(* IEC 61131-3 sources: rusty/tests/lit/single/property, 21 files *)

(* ---- called_inside_pou_where_defined.st ---- *)
// RUN: %COMPILE %s && %RUN | %CHECK %s

FUNCTION_BLOCK A
    PROPERTY_GET sayCheese: DINT
        printf('Cheese');
    END_PROPERTY

    sayCheese;
END_FUNCTION_BLOCK

FUNCTION main
    VAR
        instanceA : A;
    END_VAR

    // CHECK: Cheese
    instanceA();
END_FUNCTION

(* ---- complex.st ---- *)
// RUN: %COMPILE %s && %RUN | %CHECK %s
FUNCTION_BLOCK fb
VAR
  x : DINT;
  foo: nest_level1;
  END_VAR
END_FUNCTION_BLOCK

FUNCTION_BLOCK nest_level1
VAR
  foo: nest_level2;
END_VAR
END_FUNCTION_BLOCK

FUNCTION_BLOCK nest_level2
VAR
  foo: DINT := 0;
END_VAR
    PROPERTY_GET myProp: DINT
      myProp := foo + 5;
    END_PROPERTY

    PROPERTY_SET myProp: DINT
      foo := myProp + foo;
    END_PROPERTY
END_FUNCTION_BLOCK

FUNCTION main
    VAR
        bar: fb;
        x : DINT := 1;
    END_VAR

printf('%d$N', bar.foo.foo.myProp);   // CHECK: 5
bar.foo.foo.myProp := 10;
printf('%d$N', bar.foo.foo.myProp);   // CHECK: 15
END_FUNCTION

(* ---- get_with_early_return.st ---- *)
// RUN: %COMPILE %s && %RUN | %CHECK %s

// A RETURN in a getter returns the value of the property variable at the RETURN
FUNCTION_BLOCK fb
    VAR_INPUT
        mode : DINT;
    END_VAR

    PROPERTY_GET p : DINT
        IF mode = 1 THEN
            p := 5;
            RETURN;
        END_IF

        CASE mode OF
            2:
                p := 7;
                RETURN;
        END_CASE

        WHILE TRUE DO
            p := 8;
            IF mode = 3 THEN
                RETURN;
            END_IF
            EXIT;
        END_WHILE

        p := 6;
    END_PROPERTY
END_FUNCTION_BLOCK

FUNCTION main : DINT
    VAR
        f : fb;
    END_VAR

    // CHECK: 6
    printf('%d$N', f.p);

    f.mode := 1;
    // CHECK: 5
    printf('%d$N', f.p);

    f.mode := 2;
    // CHECK: 7
    printf('%d$N', f.p);

    f.mode := 3;
    // CHECK: 8
    printf('%d$N', f.p);
END_FUNCTION

(* ---- getter_used_in_array_indexing.st ---- *)
// RUN: %COMPILE %s && %RUN | %CHECK %s

FUNCTION_BLOCK fb
    VAR
        localVariable: ARRAY[1..5] OF DINT := [2, 4, 8, 16, 32];
    END_VAR

    PROPERTY_GET foo: ARRAY[1..5] OF DINT
        foo := localVariable;
    END_PROPERTY

    PROPERTY_GET bar: DINT
        bar := 3;
    END_PROPERTY
END_FUNCTION_BLOCK

FUNCTION main
    VAR
        instance: fb;

        arrayValue: ARRAY[1..5] OF DINT;
        arrayIndex: DINT;
    END_VAR

    printf('%d$N', instance.foo[instance.bar]); // CHECK: 8
END_FUNCTION

(* ---- modify_array_value_with_get_and_set.st ---- *)
// RUN: %COMPILE %s && %RUN | %CHECK %s

FUNCTION_BLOCK fb
    VAR
        localArray: ARRAY[1..5] OF DINT := [1, 2, 3, 4, 5];
    END_VAR

    PROPERTY_GET foo: ARRAY[1..5] OF DINT
        foo := localArray;
    END_PROPERTY

    PROPERTY_SET foo: ARRAY[1..5] OF DINT
        localArray := foo;
    END_PROPERTY
END_FUNCTION_BLOCK

FUNCTION main
    VAR
        localArray: ARRAY[1..5] OF DINT;
        fbInstance: fb;
    END_VAR

    localArray := fbInstance.foo;
    localArray[1] := 5;
    localArray[5] := 1;

    fbInstance.foo := localArray;

    printf('%d$N', fbInstance.foo[1]); // CHECK: 5
    printf('%d$N', fbInstance.foo[5]); // CHECK: 1
END_FUNCTION

(* ---- multiply_properties_single_pou.st ---- *)
// RUN: %COMPILE %s && %RUN | %CHECK %s

FUNCTION_BLOCK A
    VAR
        foo : DINT;
    END_VAR

    PROPERTY_GET increaseFooBy10: DINT
        printf('Inside increaseFooBy10$N');
        foo := foo + 10;
    END_PROPERTY

    PROPERTY_GET increaseFooBy20: DINT
        printf('Inside increaseFooBy20$N');
        foo := foo + 20;
    END_PROPERTY

    PROPERTY_GET increaseFooBy30: DINT
        printf('Inside increaseFooBy30$N');
        increaseFooBy20;
        increaseFooBy10;
    END_PROPERTY

    PROPERTY_GET readFoo: DINT
        printf('Inside readFoo$N');
        readFoo := foo;
    END_PROPERTY
END_FUNCTION_BLOCK

FUNCTION main
    VAR
        instanceA : A;
        result : DINT;
    END_VAR

    // CHECK: Inside increaseFooBy10
    instanceA.increaseFooBy10;

    // CHECK: Inside increaseFooBy20
    instanceA.increaseFooBy20;

    // CHECK: Inside increaseFooBy30
    // CHECK: Inside increaseFooBy20
    // CHECK: Inside increaseFooBy10
    instanceA.increaseFooBy30;

    // CHECK: Inside readFoo
    // CHECK: 60
    printf('%d$N', instanceA.readFoo);
END_FUNCTION

(* ---- nested.st ---- *)
// RUN: %COMPILE %s && %RUN | %CHECK %s

FUNCTION_BLOCK A
    VAR
        instanceB : B;
    END_VAR
END_FUNCTION_BLOCK

FUNCTION_BLOCK B
    VAR
        instanceC : C;
    END_VAR
END_FUNCTION_BLOCK

FUNCTION_BLOCK C
    VAR
        localPrivateVariable : DINT := 69;
    END_VAR

    PROPERTY_GET foo: DINT
        printf('Inside getter$N');
        foo := localPrivateVariable;
    END_PROPERTY

    PROPERTY_SET foo: DINT
        printf('Inside setter$N');
        localPrivateVariable := localPrivateVariable + foo;
    END_PROPERTY
END_FUNCTION_BLOCK

FUNCTION main
    VAR
        instanceA : A;
    END_VAR

    // CHECK: Inside getter
    // CHECK: 69
    printf('%d$N', instanceA.instanceB.instanceC.foo);

    // CHECK: Inside setter
    instanceA.instanceB.instanceC.foo := 351;

    // CHECK: Inside getter
    // CHECK: 420
    printf('%d$N', instanceA.instanceB.instanceC.foo);
END_FUNCTION

(* ---- oop_extended_fb_calls_property_in_another_property.st ---- *)
// RUN: %COMPILE %s && %RUN | %CHECK %s

FUNCTION_BLOCK fb
    PROPERTY_GET foo: DINT
        foo := 69;
    END_PROPERTY
END_FUNCTION_BLOCK

FUNCTION_BLOCK fb2 EXTENDS fb
    PROPERTY_GET bar: DINT
        bar := foo;
    END_PROPERTY
END_FUNCTION_BLOCK

FUNCTION main
    VAR
        fbInstance: fb2;
    END_VAR

    printf('%d$N', fbInstance.bar); // CHECK: 69
END_FUNCTION

(* ---- oop_extended_function_block.st ---- *)
// RUN: %COMPILE %s && %RUN | %CHECK %s

FUNCTION_BLOCK fb
    VAR
        returnValue: ARRAY[1..5] OF STRING := ['a', 'b', 'c', 'd', 'e'];
    END_VAR

    PROPERTY_GET foo: ARRAY[1..5] OF STRING
        foo := returnValue;
    END_PROPERTY

    PROPERTY_GET bar: DINT
        bar := 5;
    END_PROPERTY
END_FUNCTION_BLOCK

FUNCTION_BLOCK fb2 EXTENDS fb
END_FUNCTION_BLOCK

FUNCTION main
    VAR
        fbInstance: fb2;
    END_VAR

    printf('%s$N', REF(fbInstance.foo[1])); // CHECK: a
    printf('%d$N', fbInstance.bar); // CHECK: 5
END_FUNCTION

(* ---- oop_inheritance.st ---- *)
// RUN: %COMPILE %s && %RUN | %CHECK %s

INTERFACE intf
    PROPERTY_GET prop: DINT END_PROPERTY
    PROPERTY_SET prop: DINT END_PROPERTY
END_INTERFACE

FUNCTION_BLOCK fb IMPLEMENTS intf
    VAR
        localPrivateVariable: DINT := 69;
    END_VAR

    PROPERTY_GET prop: DINT
        prop := localPrivateVariable;
    END_PROPERTY

    PROPERTY_SET prop: DINT
        // This should never be called when using fb2 because it will be overridden
        localPrivateVariable := 0;
    END_PROPERTY
END_FUNCTION_BLOCK

FUNCTION_BLOCK fb2 EXTENDS fb
    PROPERTY_SET prop: DINT
        localPrivateVariable := prop;
    END_PROPERTY
END_FUNCTION_BLOCK

FUNCTION main: DINT
    VAR
        instance: fb2;
    END_VAR

    // This will call the getter from fb
    printf('%d$N', instance.prop); // CHECK: 69

    // This will call the setter from fb2
    instance.prop := 420;
    printf('%d$N', instance.prop); // CHECK: 420
END_FUNCTION

(* ---- oop_interface_extension.st ---- *)
// RUN: %COMPILE %s && %RUN | %CHECK %s

FUNCTION_BLOCK fb1
    VAR
        localPrivateVariable: DINT := 68;
    END_VAR

    PROPERTY_GET prop: DINT
        prop := localPrivateVariable;
    END_PROPERTY
END_FUNCTION_BLOCK

FUNCTION_BLOCK fb2 EXTENDS fb1
    PROPERTY_SET prop: DINT
        VAR
            x: DINT;
        END_VAR

        x := prop + 1;
        localPrivateVariable := x;
    END_PROPERTY
END_FUNCTION_BLOCK

FUNCTION main
    VAR
        instance: fb2;
    END_VAR

    instance.prop := 68;
    printf('%d$N', instance.prop); // CHECK: 69
END_FUNCTION

(* ---- oop_interface_extension_call_in_fb_body.st ---- *)
// RUN: %COMPILE %s && %RUN | %CHECK %s

FUNCTION_BLOCK fb1
    VAR
        localPrivateVariable: DINT := 67;
    END_VAR

    PROPERTY_GET prop: DINT
        prop := localPrivateVariable;
    END_PROPERTY
END_FUNCTION_BLOCK

FUNCTION_BLOCK fb2 EXTENDS fb1
    PROPERTY_SET prop: DINT
        VAR
            x: DINT;
        END_VAR

        x := prop + 1;
        localPrivateVariable := x;
    END_PROPERTY

    prop := prop + 1;
END_FUNCTION_BLOCK

FUNCTION main
    VAR
        instance: fb2;
    END_VAR

    instance();
    printf('%d$N', instance.prop); // CHECK: 69
END_FUNCTION

(* ---- property_get_with_reference_to_return_type.st ---- *)
// RUN: %COMPILE %s && %RUN | %CHECK %s
PROGRAM test
VAR
	fb	: fb;
END_VAR

printf('%d$N', fb.myStructuredVar.x);

END_PROGRAM

FUNCTION_BLOCK fb
VAR
	_myStructuredVar	: structuredTypeOrFb;
END_VAR

PROPERTY_GET myStructuredVar : REFERENCE TO structuredTypeOrFb
	myStructuredVar REF= _myStructuredVar;
END_PROPERTY

END_FUNCTION_BLOCK

TYPE structuredTypeOrFb :
	STRUCT
		x	: INT := 42;
	END_STRUCT
END_TYPE

FUNCTION main
    // CHECK: 42
    test();
END_FUNCTION

(* ---- property_get_with_referenceto_return_type_in_expression.st ---- *)
// RUN: %COMPILE %s && %RUN | %CHECK %s
PROGRAM test
VAR
	fb : fb;
    tempStruct_store : structuredTypeOrFb;
    tempStruct : REFERENCE TO structuredTypeOrFb;
    y: INT;
END_VAR

tempStruct_store.x := 51;
tempStruct REF= tempStruct_store;

// CHECK: Pre-init value: 51
printf('Pre-init value: %d$N', tempStruct.x);

fb.myStructuredVar := tempStruct;

// CHECK: Post-init value: 51
printf('Post-init value: %d$N', fb.myStructuredVar.x);

// CHECK: Expression value: 52
y := fb.myStructuredVar.x + 1;
printf('Expression value: %d$N', y);

END_PROGRAM

FUNCTION_BLOCK fb
VAR
	_myStructuredVar	: structuredTypeOrFb;
END_VAR

PROPERTY_GET myStructuredVar : REFERENCE TO structuredTypeOrFb
	myStructuredVar REF= _myStructuredVar;
END_PROPERTY

PROPERTY_SET myStructuredVar : REFERENCE TO structuredTypeOrFb
	_myStructuredVar := myStructuredVar;
END_PROPERTY

END_FUNCTION_BLOCK

TYPE structuredTypeOrFb :
	STRUCT
		x	: INT := 42;
	END_STRUCT
END_TYPE

FUNCTION main
    test();
END_FUNCTION

(* ---- property_set_with_reference_to_return_type.st ---- *)
// RUN: %COMPILE %s && %RUN | %CHECK %s
PROGRAM test
VAR
	fb : fb;
    tempStruct_store : structuredTypeOrFb;
    tempStruct : REFERENCE TO structuredTypeOrFb;
END_VAR

tempStruct_store.x := 51;
tempStruct REF= tempStruct_store;

// CHECK: Pre-init value: 51
printf('Pre-init value: %d$N', tempStruct.x);

fb.myStructuredVar := tempStruct;

// CHECK: Post-init value: 51
printf('Post-init value: %d$N', fb.myStructuredVar.x);

END_PROGRAM

FUNCTION_BLOCK fb
VAR
	_myStructuredVar	: structuredTypeOrFb;
END_VAR

PROPERTY_GET myStructuredVar : REFERENCE TO structuredTypeOrFb
	myStructuredVar REF= _myStructuredVar;
END_PROPERTY

PROPERTY_SET myStructuredVar : REFERENCE TO structuredTypeOrFb
	_myStructuredVar := myStructuredVar;
END_PROPERTY

END_FUNCTION_BLOCK

TYPE structuredTypeOrFb :
	STRUCT
		x	: INT := 42;
	END_STRUCT
END_TYPE

FUNCTION main
    test();
END_FUNCTION

(* ---- property_used_in_action.st ---- *)
// RUN: %COMPILE %s && %RUN | %CHECK %s
FUNCTION_BLOCK A
    VAR
        x : DINT := 42;
    END_VAR
    PROPERTY_GET foo: DINT
        foo := x;
    END_PROPERTY

    METHOD bar : DINT
        bar := foo;
    END_METHOD
END_FUNCTION_BLOCK

ACTIONS
    ACTION baz
        // CHECK: 42
        printf('%d$N', bar());
        // CHECK: 42
        printf('%d$N', foo);
    END_ACTION
END_ACTIONS

FUNCTION main
    VAR
        instanceA : A;
    END_VAR
        instanceA.baz();
END_FUNCTION

(* ---- property_with_chained_reference_to_return_type.st ---- *)
// RUN: %COMPILE %s && %RUN | %CHECK %s
PROGRAM test
VAR
	fb : fb;
    y : INT;
    tempStruct_store : structuredTypeOrFb;
    tempStruct2_store : structuredTypeOrFb2;
    tempStruct : REFERENCE TO structuredTypeOrFb;
END_VAR

tempStruct2_store.x := 51;
tempStruct_store.subType REF= tempStruct2_store;
tempStruct REF= tempStruct_store;

// CHECK: Pre-init value: 51
printf('Pre-init value: %d$N', tempStruct.subType.x);

fb.myStructuredVar := tempStruct;

// CHECK: Post-init value: 51
printf('Post-init value: %d$N', fb.myStructuredVar.subType.x);

END_PROGRAM

FUNCTION_BLOCK fb
VAR
	_myStructuredVar	: structuredTypeOrFb;
END_VAR

PROPERTY_GET myStructuredVar : REFERENCE TO structuredTypeOrFb
	myStructuredVar REF= _myStructuredVar;
END_PROPERTY

PROPERTY_SET myStructuredVar : REFERENCE TO structuredTypeOrFb
	_myStructuredVar := myStructuredVar;
END_PROPERTY

END_FUNCTION_BLOCK

TYPE structuredTypeOrFb :
	STRUCT
		subType : REFERENCE TO structuredTypeOrFb2;
	END_STRUCT
END_TYPE

TYPE structuredTypeOrFb2 :
	STRUCT
		x : INT := 42;
	END_STRUCT
END_TYPE

FUNCTION main
    test();
END_FUNCTION

(* ---- property_with_local_variables.st ---- *)
// RUN: %COMPILE %s && %RUN | %CHECK %s
FUNCTION_BLOCK fb
    VAR
        localPrivateVariable: DINT := 5;
    END_VAR

    PROPERTY_GET foo: DINT
        VAR
            one: DINT := 1;
        END_VAR

        foo := localPrivateVariable + one;
    END_PROPERTY

    PROPERTY_SET foo: DINT
        VAR
            two: DINT := 2;
            three: DINT := 3;
        END_VAR
        localPrivateVariable := two + foo + three;
    END_PROPERTY
END_FUNCTION_BLOCK

FUNCTION main
    VAR
        localVariable: DINT;
        instance: fb;
    END_VAR

    // Retrieving the getter return value using another variable
    localVariable := instance.foo;
    printf('%d$N', localVariable); // CHECK: 6

    // Retrieving the getter return value using the property directly
    printf('%d$N', instance.foo); // CHECK: 6

    instance.foo := 10;
    printf('%d$N', instance.foo); // CHECK: 16
END_FUNCTION

(* ---- same_property_in_different_pous_called_in_method.st ---- *)
// RUN: %COMPILE %s && %RUN | %CHECK %s
FUNCTION_BLOCK A
    VAR
        x : DINT := 42;
    END_VAR

    PROPERTY_GET foo: DINT
        foo := x;
    END_PROPERTY
END_FUNCTION_BLOCK

FUNCTION_BLOCK B
    VAR
        x : DINT := 69;
    END_VAR

    PROPERTY_GET foo: DINT
        foo := x;
    END_PROPERTY

    METHOD bar : DINT
    VAR
        instanceA : A;
    END_VAR
        bar := foo;
    END_METHOD

    METHOD baz : DINT
    VAR
        instanceA : A;
    END_VAR
        baz := instanceA.foo;
    END_METHOD
END_FUNCTION_BLOCK

FUNCTION main
    VAR
        instanceB : B;
    END_VAR

    printf('%d$N', instanceB.bar()); // CHECK: 69
    printf('%d$N', instanceB.baz()); // CHECK: 42
END_FUNCTION

(* ---- simple.st ---- *)
// RUN: %COMPILE %s && %RUN | %CHECK %s
FUNCTION_BLOCK fb
    VAR
        localPrivateVariable : DINT := 5;
    END_VAR

    PROPERTY_GET foo: DINT
        foo := localPrivateVariable;
    END_PROPERTY

    PROPERTY_SET foo: DINT
        localPrivateVariable := foo + 5;
    END_PROPERTY
END_FUNCTION_BLOCK

FUNCTION main
    VAR
        localVariable : DINT;
        instance : fb;
    END_VAR

    // Retrieving the getter return value using another variable
    localVariable := instance.foo;
    printf('%d$N', localVariable);  // CHECK: 5

    // Retrieving the getter return value using the property directly
    printf('%d$N', instance.foo);   // CHECK: 5

    instance.foo := 10;
    printf('%d$N', instance.foo);   // CHECK: 15
END_FUNCTION

(* ---- struct_return_type.st ---- *)
// RUN: %COMPILE %s && %RUN | %CHECK %s

TYPE
    Transaction: STRUCT
        id: DINT;
        values: ARRAY[1..10] OF DINT;
    END_STRUCT
END_TYPE

FUNCTION print_txn
    VAR_INPUT {ref}
        value: Transaction;
    END_VAR

    VAR
        idx: DINT;
    END_VAR

    printf('{ id: %d, values: [', value.id);
    FOR idx := 1 TO 10 DO
        IF idx > 1 THEN
            printf(', ');
        END_IF;
        printf('%d', value.values[idx]);
    END_FOR;
    printf('] }$N');
END_FUNCTION

FUNCTION_BLOCK fb
    VAR
        localPrivateVariable: DINT := 5;
        returnValue: Transaction;
    END_VAR

    PROPERTY_GET foo: Transaction
        printf('Inside getter$N');

        // Uninitialized
        IF returnValue.id = 0 THEN
            returnValue.id := 1;
            returnValue.values := [1, 2, 4, 8, 16, 32, 64, 128, 256, 512];
        END_IF

        foo := returnValue;
    END_PROPERTY

    PROPERTY_SET foo: Transaction
        printf('Inside setter$N');

        returnValue := foo;
    END_PROPERTY
END_FUNCTION_BLOCK

FUNCTION main
    VAR
        instance: fb;
        localTransaction: Transaction;
    END_VAR

    // CHECK: Inside getter
    // CHECK: { id: 1, values: [1, 2, 4, 8, 16, 32, 64, 128, 256, 512] }
    print_txn(instance.foo);

    // CHECK: Inside getter
    // CHECK: Inside setter
    // CHECK: Inside getter
    // CHECK: { id: 69, values: [1, 2, 4, 8, 16, 32, 64, 128, 256, 512] }
    localTransaction := instance.foo;
    localTransaction.id := 69;
    instance.foo := localTransaction;
    print_txn(instance.foo);
END_FUNCTION
